// TIA Portal V21 export
// export: Created 2026-11-10T19:16:53.6419853Z, ExportSetting WithDefaults, DisplayName Totally Integrated Automation Portal, DisplayVersion V21 Update 3, DisplayName STEP 7 Professional, DisplayVersion V21 Update 3, DisplayName STEP 7 Safety, DisplayVersion V21, DisplayName Tech WebApplication, DisplayVersion V21, DisplayName WinCC Basic/Comfort/Advanced, DisplayVersion V21 Update 3, DisplayName WinCC Unified, DisplayVersion V21 Update 3
TYPE "UDT_Inner"
// stored: IsFailsafeCompliant false
   STRUCT
      Temp : Real := 21.5;
      Input { ExternalWritable := 'False'} : Bool;
      Static { S7_SetPoint := 'True'} : Int := 3;
      "Return" { ExternalAccessible := 'False'; ExternalVisible := 'False'; ExternalWritable := 'False'} : DInt;
      Arr { ExternalVisible := 'False'} : Array[1..3] of Int;
   END_STRUCT;
END_TYPE
